(* IEC 61131-3 sources: axsharp/src/ix.templates/working/templates/ixblazor/ax/src, 3 files *)

(* ---- counter_oop.st ---- *)
{#ix-attr:[Container(Layout.Wrap)]}
CLASS PUBLIC counter_oop
    VAR PUBLIC
        Counter : ULINT;
        AllowCounter : BOOL;
    END_VAR

    METHOD PUBLIC RunCounter
        IF (AllowCounter) THEN
            Counter := Counter + ULINT#1;
        END_IF;
    END_METHOD

END_CLASS

(* ---- configuration.st ---- *)
CONFIGURATION MyConfiguration
    TASK Main(Interval := T#10ms, Priority := 1);
    PROGRAM P1 WITH Main: MyProgram;

    VAR_GLOBAL
        oop_counter : counter_oop;
    END_VAR
END_CONFIGURATION

(* ---- program.st ---- *)
PROGRAM MyProgram
    VAR_EXTERNAL
        oop_counter : counter_oop;
    END_VAR
    oop_counter.RunCounter();
END_PROGRAM
